FUNCTION_BLOCK basicSensorGenerico (* Logica unica do sensor generico (4-20 mA ou comunicacao) *)
  (* Standard: 61499-2 *)
  (* Version 2.2, 12/11/2026, Hidryco, Hidryco, 2.2: aviso e erro do proprio dispositivo por comunicacao (fldAvisoDisp/fldErroDisp, REQ_FB_DISP): erro diferente de 0 = falha do sensor (cfgTempoFalha); aviso = alarme almAviso; codigos stsCodigoErro/stsCodigoAviso para o diagnostico. 2.1: cfgSkid = sensor sempre habilitado. 2.0: falha do 4-20 mA abaixo de 3800 ou acima de 22000 (eram 3600/21000), confirmada em cfgTempoFalha. 1.9: stsAtivoHH/stsAtivoH (alarme com o tempo do alarme e sem memoria; some quando o valor volta) e stsDisponivel (sensor habilitado, com leitura e sem falha) no CNF. 1.8: limites dos alarmes em unidade de engenharia para o grafico da IHM (stsLimHH..LL; nivel: % x altura maxima / 100). 1.7: stsFalhaSensor (STS_FALHA_SENSOR) so com a falha do sensor (fora da faixa ou falha do instrumento), sem a comunicacao; stsFalhaAtiva e o alarme de falha com qualquer falha. 1.6: IHM: valor, % e bruto no maximo 1 vez por segundo (evento TICK de 1 s); estado, falha e alarmes na hora. 1.5: saida stsFalhaComunicacao (comunicacao do instrumento ou conexao Modbus offline). 1.4: stsFalhaSensor (STS_FALHA_SENSOR na IHM) = falha ativa: sensor em falha agora, sem memoria nem reset; o alarme de falha segue. 1.3: sensor de nivel (cfgNivel) compara os alarmes HH/H/L/LL com a % da altura maxima (setpoints em %); os demais com o valor. 1.2: falha do sinal tambem pelo status da conexao Modbus (fldConexao INT, 1 = online) com cfgUsaConexao, nos dois modos (4-20 mA lido por remota e comunicacao). 1.1: inibicao de L/LL pelo processo e condicao instantanea de cada limite. 1.0: padrao SE.App2CommonProcess - escala, falha NAMUR confirmada por tempo, alarmes HH/H/L/LL com tempo proprio e memoria ate o reset, supressao em falha *)
  PACKAGE Hidryco.HidrycoLib;
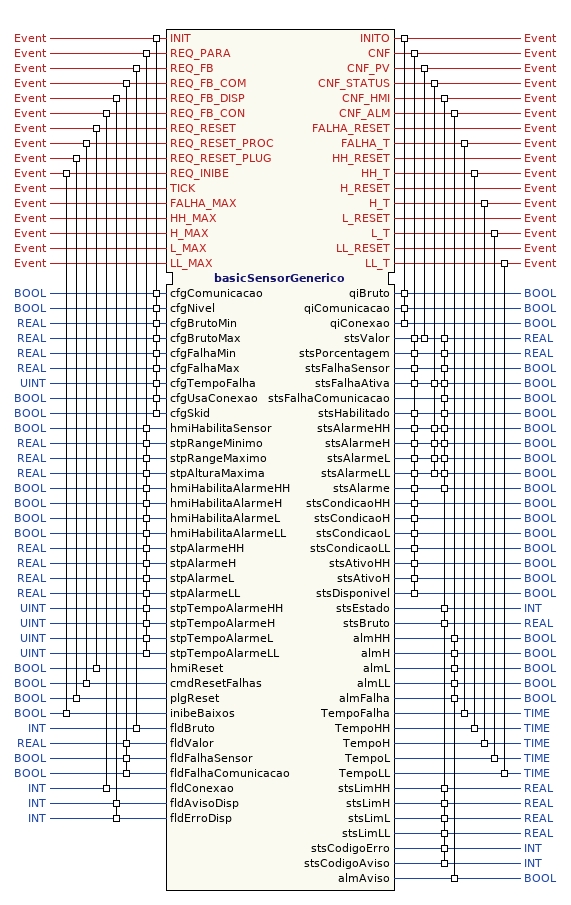
  EVENT_INPUT
    INIT WITH cfgComunicacao, cfgNivel, cfgBrutoMin, cfgBrutoMax, cfgFalhaMin, cfgFalhaMax, cfgTempoFalha, cfgUsaConexao, cfgSkid; (* Inicializacao *)
    REQ_PARA WITH hmiHabilitaSensor, stpRangeMinimo, stpRangeMaximo, stpAlturaMaxima, hmiHabilitaAlarmeHH, hmiHabilitaAlarmeH, hmiHabilitaAlarmeL, hmiHabilitaAlarmeLL, stpAlarmeHH, stpAlarmeH, stpAlarmeL, stpAlarmeLL, stpTempoAlarmeHH, stpTempoAlarmeH, stpTempoAlarmeL, stpTempoAlarmeLL; (* Parametros da IHM (persistentes) *)
    REQ_FB WITH fldBruto; (* Leitura 4-20 mA *)
    REQ_FB_COM WITH fldValor, fldFalhaSensor, fldFalhaComunicacao; (* Leitura por comunicacao *)
    REQ_FB_DISP WITH fldAvisoDisp, fldErroDisp; (* Aviso e erro do proprio dispositivo (comunicacao) *)
    REQ_FB_CON WITH fldConexao; (* Status da conexao Modbus (comunicacao) *)
    REQ_RESET WITH hmiReset; (* Reset pela IHM *)
    REQ_RESET_PROC WITH cmdResetFalhas; (* Reset pelo processo *)
    REQ_RESET_PLUG WITH plgReset; (* Reset pelo plug ISensorStatus *)
    REQ_INIBE WITH inibeBaixos; (* Inibicao dos alarmes L e LL pelo processo *)
    TICK; (* Base de 1 s para atualizar a IHM *)
    FALHA_MAX; (* Fim do tempo de confirmacao da falha (E_DELAY) *)
    HH_MAX; (* Fim do tempo do alarme HH (E_DELAY) *)
    H_MAX; (* Fim do tempo do alarme H (E_DELAY) *)
    L_MAX; (* Fim do tempo do alarme L (E_DELAY) *)
    LL_MAX; (* Fim do tempo do alarme LL (E_DELAY) *)
  END_EVENT
  EVENT_OUTPUT
    INITO WITH qiBruto, qiComunicacao, qiConexao; (* Inicializacao concluida *)
    CNF WITH stsValor, stsPorcentagem, stsFalhaSensor, stsFalhaAtiva, stsHabilitado, stsAlarmeHH, stsAlarmeH, stsAlarmeL, stsAlarmeLL, stsAlarme, stsCondicaoHH, stsCondicaoH, stsCondicaoL, stsCondicaoLL, stsAtivoHH, stsAtivoH, stsDisponivel; (* Status para o processo (na mudanca) *)
    CNF_PV WITH stsValor; (* Valor para o plug (na mudanca) *)
    CNF_STATUS WITH stsAlarmeHH, stsAlarmeH, stsAlarmeL, stsAlarmeLL, stsFalhaAtiva; (* Alarmes para o plug (na mudanca) *)
    CNF_HMI WITH stsValor, stsPorcentagem, stsEstado, stsFalhaSensor, stsFalhaAtiva, stsHabilitado, stsAlarmeHH, stsAlarmeH, stsAlarmeL, stsAlarmeLL, stsAlarme, stsBruto, stsFalhaComunicacao, stsLimHH, stsLimH, stsLimL, stsLimLL, stsCodigoErro, stsCodigoAviso; (* Status para a IHM (na mudanca) *)
    CNF_ALM WITH almHH, almH, almL, almLL, almFalha, almAviso; (* Alarmes para os ALARM_BIT (na mudanca) *)
    FALHA_RESET; (* Cancela o tempo de falha (E_DELAY.STOP) - sai antes do FALHA_T *)
    FALHA_T WITH TempoFalha; (* Inicia o tempo de falha (E_DELAY.START) *)
    HH_RESET; (* Cancela o tempo do alarme HH - sai antes do HH_T *)
    HH_T WITH TempoHH; (* Inicia o tempo do alarme HH *)
    H_RESET; (* Cancela o tempo do alarme H - sai antes do H_T *)
    H_T WITH TempoH; (* Inicia o tempo do alarme H *)
    L_RESET; (* Cancela o tempo do alarme L - sai antes do L_T *)
    L_T WITH TempoL; (* Inicia o tempo do alarme L *)
    LL_RESET; (* Cancela o tempo do alarme LL - sai antes do LL_T *)
    LL_T WITH TempoLL; (* Inicia o tempo do alarme LL *)
  END_EVENT
  VAR_INPUT
    cfgComunicacao : BOOL := FALSE; (* FALSE = entrada 4-20 mA (stsSensorBruto), TRUE = valor por comunicacao (stsEntrada, ja em unidade de engenharia) *)
    cfgNivel : BOOL := FALSE; (* TRUE = sensor de nivel: calcula % sobre a altura maxima *)
    cfgBrutoMin : REAL := 4000.0; (* Valor bruto em 4 mA (TM3: 4000) *)
    cfgBrutoMax : REAL := 20000.0; (* Valor bruto em 20 mA (TM3: 20000) *)
    cfgFalhaMin : REAL := 3800.0; (* Abaixo deste bruto = falha (3,8 mA) *)
    cfgFalhaMax : REAL := 22000.0; (* Acima deste bruto = falha (22,0 mA) *)
    cfgTempoFalha : UINT := 5; (* Tempo para confirmar a falha do sinal (s) *)
    cfgUsaConexao : BOOL := FALSE; (* TRUE = sinal em falha tambem quando o status da conexao Modbus (stsConexao, INT) for diferente de 1 (4-20 mA por remota ou comunicacao) *)
    cfgSkid : BOOL := FALSE; (* TRUE = valor de skid (ja escalado no equipamento): sensor sempre habilitado, sem ajustes na IHM *)
    hmiHabilitaSensor : BOOL; (* IHM: sensor habilitado *)
    stpRangeMinimo : REAL; (* IHM: valor de engenharia em 4 mA *)
    stpRangeMaximo : REAL; (* IHM: valor de engenharia em 20 mA *)
    stpAlturaMaxima : REAL; (* IHM: altura maxima do tanque (nivel) *)
    hmiHabilitaAlarmeHH : BOOL; (* IHM: alarme HH habilitado *)
    hmiHabilitaAlarmeH : BOOL; (* IHM: alarme H habilitado *)
    hmiHabilitaAlarmeL : BOOL; (* IHM: alarme L habilitado *)
    hmiHabilitaAlarmeLL : BOOL; (* IHM: alarme LL habilitado *)
    stpAlarmeHH : REAL; (* IHM: setpoint do alarme HH *)
    stpAlarmeH : REAL; (* IHM: setpoint do alarme H *)
    stpAlarmeL : REAL; (* IHM: setpoint do alarme L *)
    stpAlarmeLL : REAL; (* IHM: setpoint do alarme LL *)
    stpTempoAlarmeHH : UINT; (* IHM: tempo do alarme HH (s) *)
    stpTempoAlarmeH : UINT; (* IHM: tempo do alarme H (s) *)
    stpTempoAlarmeL : UINT; (* IHM: tempo do alarme L (s) *)
    stpTempoAlarmeLL : UINT; (* IHM: tempo do alarme LL (s) *)
    hmiReset : BOOL; (* IHM: reset *)
    cmdResetFalhas : BOOL; (* Processo: reset (com E_RESET_FALHAS) *)
    plgReset : BOOL; (* Plug ISensorStatus: cmdReset *)
    inibeBaixos : BOOL; (* Processo: inibe os alarmes L e LL (ex.: pressao de recalque com as bombas paradas) *)
    fldBruto : INT; (* Campo: valor bruto 4-20 mA *)
    fldValor : REAL; (* Campo (comunicacao): valor em unidade de engenharia *)
    fldFalhaSensor : BOOL; (* Campo (comunicacao): falha do instrumento *)
    fldFalhaComunicacao : BOOL; (* Campo (comunicacao): falha de comunicacao *)
    fldConexao : INT; (* Campo (comunicacao): status da conexao Modbus (connStatusInt: 1 = online, 0 = offline) *)
    fldAvisoDisp : INT; (* Campo (comunicacao): condicao de aviso do proprio dispositivo (0 = nenhum) *)
    fldErroDisp : INT; (* Campo (comunicacao): condicao de erro do proprio dispositivo (0 = nenhum) *)
  END_VAR
  VAR_OUTPUT
    qiBruto : BOOL; (* Assina o symlink 4-20 mA (NOT cfgComunicacao) *)
    qiComunicacao : BOOL; (* Assina os symlinks de comunicacao (cfgComunicacao) *)
    qiConexao : BOOL; (* Assina o symlink do status da conexao (cfgUsaConexao) *)
    stsValor : REAL; (* Valor em unidade de engenharia (0 em falha ou desabilitado) *)
    stsPorcentagem : REAL; (* Nivel em % da altura maxima (so cfgNivel) *)
    stsFalhaSensor : BOOL; (* Falha do sensor (4-20 mA fora da faixa ou falha do instrumento), confirmada e ativa, sem a falha de comunicacao *)
    stsFalhaAtiva : BOOL; (* Qualquer falha confirmada e ativa (sensor ou comunicacao) *)
    stsFalhaComunicacao : BOOL; (* Falha de comunicacao do sensor (falha do instrumento por comunicacao ou conexao Modbus offline) *)
    stsHabilitado : BOOL; (* Sensor habilitado *)
    stsAlarmeHH : BOOL; (* Alarme HH (memorizado ate o reset; suprimido com o sinal em falha) *)
    stsAlarmeH : BOOL; (* Alarme H (memorizado ate o reset; suprimido com o sinal em falha) *)
    stsAlarmeL : BOOL; (* Alarme L (memorizado ate o reset; suprimido com o sinal em falha) *)
    stsAlarmeLL : BOOL; (* Alarme LL (memorizado ate o reset; suprimido com o sinal em falha) *)
    stsAlarme : BOOL; (* Algum alarme ativo *)
    stsCondicaoHH : BOOL; (* Valor alem do setpoint HH agora (sem tempo e sem memoria; so com o alarme habilitado e o sinal bom) *)
    stsCondicaoH : BOOL; (* Valor alem do setpoint H agora (sem tempo e sem memoria; so com o alarme habilitado e o sinal bom) *)
    stsCondicaoL : BOOL; (* Valor alem do setpoint L agora (sem tempo e sem memoria; so com o alarme habilitado e o sinal bom) *)
    stsCondicaoLL : BOOL; (* Valor alem do setpoint LL agora (sem tempo e sem memoria; so com o alarme habilitado e o sinal bom) *)
    stsAtivoHH : BOOL; (* Alarme HH com o tempo do alarme e sem memoria (some quando o valor volta; so com o alarme habilitado e o sinal bom) *)
    stsAtivoH : BOOL; (* Alarme H com o tempo do alarme e sem memoria (some quando o valor volta; so com o alarme habilitado e o sinal bom) *)
    stsDisponivel : BOOL; (* Sensor habilitado, com leitura e sem falha *)
    stsEstado : INT; (* IHM: 0 normal, 1 alerta (H/L), 2 alarme (HH/LL), 3 falha, 4 desabilitado *)
    stsBruto : REAL; (* IHM: valor bruto lido (diagnostico) *)
    almHH : BOOL; (* Entrada do ALARM_BIT HH *)
    almH : BOOL; (* Entrada do ALARM_BIT H *)
    almL : BOOL; (* Entrada do ALARM_BIT L *)
    almLL : BOOL; (* Entrada do ALARM_BIT LL *)
    almFalha : BOOL; (* Entrada do ALARM_BIT de falha do sensor *)
    TempoFalha : TIME; (* E_DELAY da falha *)
    TempoHH : TIME; (* E_DELAY do alarme HH *)
    TempoH : TIME; (* E_DELAY do alarme H *)
    TempoL : TIME; (* E_DELAY do alarme L *)
    TempoLL : TIME; (* E_DELAY do alarme LL *)
    stsLimHH : REAL; (* Limite do alarme HH em unidade de engenharia (para o grafico) *)
    stsLimH : REAL; (* Limite do alarme H em unidade de engenharia (para o grafico) *)
    stsLimL : REAL; (* Limite do alarme L em unidade de engenharia (para o grafico) *)
    stsLimLL : REAL; (* Limite do alarme LL em unidade de engenharia (para o grafico) *)
    stsCodigoErro : INT; (* IHM: codigo de erro do proprio dispositivo (0 = nenhum; diferente de 0 = falha do sensor) *)
    stsCodigoAviso : INT; (* IHM: codigo de aviso do proprio dispositivo (0 = nenhum; so alarme) *)
    almAviso : BOOL; (* Entrada do ALARM_BIT de aviso do proprio dispositivo *)
  END_VAR
  VAR
    initDone : BOOL;
    initPass : BOOL;
    fbRecebido : BOOL; (* Ja houve leitura do campo *)
    bReset : BOOL;
    bRuimAgora : BOOL; (* Sinal fora da faixa / falha agora *)
    bSensorRuim : BOOL; (* Falha do proprio sensor agora (fora da faixa 4-20 mA ou falha do instrumento), sem a comunicacao *)
    bSuprimido : BOOL; (* Alarmes suprimidos *)
    rBruto : REAL;
    rFaixa : REAL;
    rMin : REAL;
    rMax : REAL;
    bTimFalha : BOOL;
    oldTimFalha : BOOL;
    bCondHH : BOOL;
    bMemHH : BOOL;
    bTimHH : BOOL;
    oldTimHH : BOOL;
    bAcimaHH : BOOL;
    bCondH : BOOL;
    bMemH : BOOL;
    bTimH : BOOL;
    oldTimH : BOOL;
    bTempoHH : BOOL; (* Tempo do HH venceu com a condicao presente (sem memoria) *)
    bTempoH : BOOL; (* Tempo do H venceu com a condicao presente (sem memoria) *)
    bAcimaH : BOOL;
    bCondL : BOOL;
    bMemL : BOOL;
    bTimL : BOOL;
    oldTimL : BOOL;
    bAcimaL : BOOL;
    bCondLL : BOOL;
    bMemLL : BOOL;
    bTimLL : BOOL;
    oldTimLL : BOOL;
    bAcimaLL : BOOL;
    oldValor : REAL;
    oldPct : REAL;
    oldBruto : REAL;
    wSts : WORD;
    oldSts : WORD := 16#FFFF;
    wAlm : WORD;
    oldAlm : WORD := 16#FFFF;
    oldCodErro : INT := -1;
    oldCodAviso : INT := -1;
    oldEstado : INT := -1;
    hmiBruto : REAL := -1.0;
    hmiPct : REAL := -1.0;
    hmiValor : REAL := -1.0;
    rCmp : REAL; (* Valor comparado com os alarmes: % (sensor de nivel) ou valor *)
    rEscLim : REAL;
    ostsLimHH : REAL := -1.0;
    ostsLimH : REAL := -1.0;
    ostsLimL : REAL := -1.0;
    ostsLimLL : REAL := -1.0;
  END_VAR
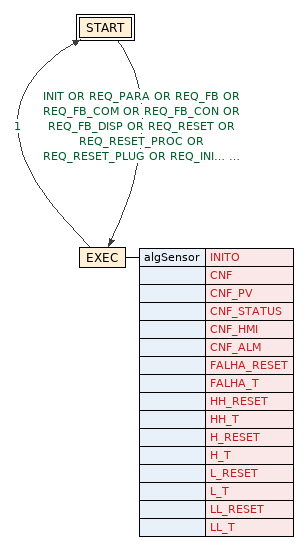
  EC_STATES
    START; (* Estado inicial *)
    EXEC : algSensor -> INITO, -> CNF, -> CNF_PV, -> CNF_STATUS, -> CNF_HMI, -> CNF_ALM, -> FALHA_RESET, -> FALHA_T, -> HH_RESET, -> HH_T, -> H_RESET, -> H_T, -> L_RESET, -> L_T, -> LL_RESET, -> LL_T; (* Executa a logica; o algoritmo decide quais eventos saem *)
  END_STATES
  EC_TRANSITIONS
    START TO EXEC := INIT OR REQ_PARA OR REQ_FB OR REQ_FB_COM OR REQ_FB_CON OR REQ_FB_DISP OR REQ_RESET OR REQ_RESET_PROC OR REQ_RESET_PLUG OR REQ_INIBE OR FALHA_MAX OR HH_MAX OR H_MAX OR L_MAX OR LL_MAX OR TICK;
    EXEC TO START := 1;
  END_TRANSITIONS
  ALGORITHM algSensor IN ST: (* Logica completa do sensor (um unico algoritmo) *)
(* =====================================================================
   basicSensorGenerico v1.1 - logica do CAT Sensor_Generico (HidrycoLib)
   Padrao das bibliotecas Schneider (SE.App2CommonProcess):
   - eventos de saida desligados no inicio e ligados so na mudanca;
   - tempos por E_DELAY externo (X_T / X_RESET / X_MAX), um por alarme;
   - alarmes para o sistema de alarmes do EAE por ALARM_BIT (no CAT).
   Regras (definidas pelo usuario):
   - origem 4-20 mA (escala bruta e limites NAMUR offline) ou comunicacao
     (valor ja em unidade de engenharia);
   - falha do sinal confirmada apos cfgTempoFalha: valor vai a 0 e os
     alarmes ficam suprimidos; a falha vale enquanto o sinal estiver ruim, e o
     sensor volta a funcionar assim que o sinal volta;
   - durante a confirmacao o valor fica congelado (nao vai a 0 por um pico);
   - alarmes HH/H/L/LL sem histerese, cada um com o proprio tempo,
     memorizados ate o reset (IHM, processo ou plug);
   - sensor desabilitado: valor 0, sem falha e sem alarmes.
   v1.3: sensor de nivel (cfgNivel): HH/H/L/LL comparados com a % da altura maxima.
   v1.1: inibeBaixos (processo) inibe L/LL e libera a memoria deles;
         stsCondicaoX = valor alem do setpoint X agora (sem tempo, sem memoria).
   ===================================================================== *)

(* ---- 0. Eventos de saida: so sai o que for ligado abaixo ---- *)
INITO       := FALSE;
CNF         := FALSE;
CNF_PV      := FALSE;
CNF_STATUS  := FALSE;
CNF_HMI     := FALSE;
CNF_ALM     := FALSE;
FALHA_RESET := FALSE;
FALHA_T     := FALSE;
HH_RESET := FALSE; HH_T := FALSE;
H_RESET  := FALSE; H_T  := FALSE;
L_RESET  := FALSE; L_T  := FALSE;
LL_RESET := FALSE; LL_T := FALSE;

IF REQ_FB OR REQ_FB_COM OR REQ_FB_CON THEN
    fbRecebido := TRUE;                    (* campo valido a partir da 1a leitura *)
END_IF;

(* ---- 1. Inicializacao ---- *)
IF INIT THEN
    qiBruto       := NOT cfgComunicacao;   (* so assina o symlink da origem configurada *)
    qiComunicacao := cfgComunicacao;
    qiConexao     := cfgUsaConexao;           (* status da conexao: vale para 4-20 mA lido por remota e para comunicacao *)
    initDone := TRUE;
    initPass := TRUE;
    INITO    := TRUE;
END_IF;
IF NOT initDone THEN
    RETURN;
END_IF;
(* sensor de skid: nao pode ser desabilitado (vale mesmo com FALSE gravado de antes) *)
IF cfgSkid THEN
    hmiHabilitaSensor := TRUE;
END_IF;

(* ---- 2. Sinal ---- *)
IF cfgComunicacao THEN
    rBruto     := fldValor;
    bRuimAgora := fbRecebido AND (fldFalhaSensor OR fldFalhaComunicacao OR (cfgUsaConexao AND fldConexao <> 1));
    bSensorRuim := fbRecebido AND fldFalhaSensor;
ELSE
    rBruto     := INT_TO_REAL(fldBruto);
    bRuimAgora := fbRecebido AND ((rBruto < cfgFalhaMin) OR (rBruto > cfgFalhaMax) OR (cfgUsaConexao AND fldConexao <> 1));
    bSensorRuim := fbRecebido AND ((rBruto < cfgFalhaMin) OR (rBruto > cfgFalhaMax));
END_IF;

(* erro do proprio dispositivo (ex.: SC4500 por Modbus): falha do sensor, confirmada pelo mesmo tempo *)
IF fbRecebido AND (fldErroDisp <> 0) THEN
    bRuimAgora  := TRUE;
    bSensorRuim := TRUE;
END_IF;

(* ---- 3. Falha do sensor: confirmada pelo tempo; vale enquanto o sensor estiver em falha (sem memoria) ---- *)
bReset := (REQ_RESET AND hmiReset) OR (REQ_RESET_PROC AND cmdResetFalhas) OR (REQ_RESET_PLUG AND plgReset);
IF NOT hmiHabilitaSensor THEN
    stsFalhaAtiva := FALSE;
ELSE
    IF FALHA_MAX AND bRuimAgora THEN
        stsFalhaAtiva := TRUE;             (* falha confirmada *)
    END_IF;
    IF NOT bRuimAgora THEN
        stsFalhaAtiva := FALSE;            (* sinal voltou: a falha sai sozinha, sem reset *)
    END_IF;
END_IF;
(* falha de comunicacao (imediata; o tempo de deteccao e o do proprio Modbus) *)
stsFalhaComunicacao := hmiHabilitaSensor AND fbRecebido AND
    ((cfgComunicacao AND fldFalhaComunicacao) OR (cfgUsaConexao AND fldConexao <> 1));
(* STS_FALHA_SENSOR = so a falha do sensor (confirmada pelo tempo); com a comunicacao em falha o valor lido nao vale, entao nao conta *)
stsFalhaSensor := stsFalhaAtiva AND bSensorRuim AND NOT stsFalhaComunicacao;
bTimFalha := hmiHabilitaSensor AND bRuimAgora AND NOT stsFalhaAtiva;
IF bTimFalha <> oldTimFalha THEN
    IF bTimFalha THEN
        TempoFalha := TO_TIME(UINT_TO_DINT(cfgTempoFalha) * 1000);
        FALHA_T := TRUE;
    ELSE
        FALHA_RESET := TRUE;
    END_IF;
    oldTimFalha := bTimFalha;
END_IF;

(* ---- 4. Valor em unidade de engenharia ---- *)
IF NOT hmiHabilitaSensor OR NOT fbRecebido OR stsFalhaAtiva THEN
    stsValor := 0.0;                       (* desabilitado, sem leitura ou falha confirmada *)
ELSIF bRuimAgora THEN
    ;                                      (* confirmando a falha: valor congelado *)
ELSIF cfgComunicacao THEN
    stsValor := fldValor;                  (* ja chega em unidade de engenharia *)
ELSE
    rFaixa := cfgBrutoMax - cfgBrutoMin;
    IF rFaixa <> 0.0 THEN
        stsValor := stpRangeMinimo + (rBruto - cfgBrutoMin) * (stpRangeMaximo - stpRangeMinimo) / rFaixa;
        rMin := MIN(stpRangeMinimo, stpRangeMaximo);
        rMax := MAX(stpRangeMinimo, stpRangeMaximo);
        stsValor := LIMIT(rMin, stsValor, rMax);
    ELSE
        stsValor := 0.0;                   (* escala bruta invalida *)
    END_IF;
END_IF;
IF cfgNivel AND stpAlturaMaxima > 0.0 THEN
    stsPorcentagem := stsValor * 100.0 / stpAlturaMaxima;
ELSE
    stsPorcentagem := 0.0;
END_IF;
stsBruto := rBruto;
(* alarmes do sensor de nivel pela % da altura maxima; os demais pelo valor em unidade de engenharia *)
IF cfgNivel THEN
    rCmp := stsPorcentagem;
ELSE
    rCmp := stsValor;
END_IF;

(* ---- 5. Alarmes (suprimidos com o sensor desabilitado, sem leitura ou em falha) ---- *)
bSuprimido := NOT hmiHabilitaSensor OR NOT fbRecebido OR bRuimAgora OR stsFalhaAtiva;
bAcimaHH := rCmp > stpAlarmeHH;
bCondHH := hmiHabilitaAlarmeHH AND NOT bSuprimido AND bAcimaHH;
stsCondicaoHH := bCondHH;
IF HH_MAX AND bCondHH THEN
    bTempoHH := TRUE;                     (* com tempo, sem memoria *)
    bMemHH := TRUE;                       (* tempo do alarme HH venceu com a condicao presente *)
END_IF;
IF bReset AND NOT bCondHH THEN
    bMemHH := FALSE;                      (* reset so libera se a condicao ja sumiu *)
END_IF;
IF NOT hmiHabilitaAlarmeHH OR NOT hmiHabilitaSensor THEN
    bMemHH := FALSE;                      (* alarme ou sensor desabilitado zera o alarme *)
END_IF;
IF NOT bCondHH THEN
    bTempoHH := FALSE;                    (* condicao sumiu: sai na hora *)
END_IF;
(* o tempo conta a cada vez que a condicao aparece, mesmo com o alarme ainda memorizado (para o stsAtivoHH) *)
bTimHH := bCondHH AND NOT bTempoHH;
IF bTimHH <> oldTimHH THEN
    IF bTimHH THEN
        TempoHH := TO_TIME(UINT_TO_DINT(stpTempoAlarmeHH) * 1000);
        HH_T := TRUE;
    ELSE
        HH_RESET := TRUE;
    END_IF;
    oldTimHH := bTimHH;
END_IF;
stsAlarmeHH := bMemHH AND NOT bSuprimido;
stsAtivoHH := bTempoHH AND bCondHH;

bAcimaH := rCmp > stpAlarmeH;
bCondH := hmiHabilitaAlarmeH AND NOT bSuprimido AND bAcimaH;
stsCondicaoH := bCondH;
IF H_MAX AND bCondH THEN
    bTempoH := TRUE;                     (* com tempo, sem memoria *)
    bMemH := TRUE;                       (* tempo do alarme H venceu com a condicao presente *)
END_IF;
IF bReset AND NOT bCondH THEN
    bMemH := FALSE;                      (* reset so libera se a condicao ja sumiu *)
END_IF;
IF NOT hmiHabilitaAlarmeH OR NOT hmiHabilitaSensor THEN
    bMemH := FALSE;                      (* alarme ou sensor desabilitado zera o alarme *)
END_IF;
IF NOT bCondH THEN
    bTempoH := FALSE;                    (* condicao sumiu: sai na hora *)
END_IF;
(* o tempo conta a cada vez que a condicao aparece, mesmo com o alarme ainda memorizado (para o stsAtivoH) *)
bTimH := bCondH AND NOT bTempoH;
IF bTimH <> oldTimH THEN
    IF bTimH THEN
        TempoH := TO_TIME(UINT_TO_DINT(stpTempoAlarmeH) * 1000);
        H_T := TRUE;
    ELSE
        H_RESET := TRUE;
    END_IF;
    oldTimH := bTimH;
END_IF;
stsAlarmeH := bMemH AND NOT bSuprimido;
stsAtivoH := bTempoH AND bCondH;

bAcimaL := rCmp < stpAlarmeL;
bCondL := hmiHabilitaAlarmeL AND NOT bSuprimido AND bAcimaL AND NOT inibeBaixos;
stsCondicaoL := bCondL;
IF inibeBaixos THEN
    bMemL := FALSE;                      (* inibido pelo processo: libera o que estava memorizado *)
END_IF;
IF L_MAX AND bCondL THEN
    bMemL := TRUE;                       (* tempo do alarme L venceu com a condicao presente *)
END_IF;
IF bReset AND NOT bCondL THEN
    bMemL := FALSE;                      (* reset so libera se a condicao ja sumiu *)
END_IF;
IF NOT hmiHabilitaAlarmeL OR NOT hmiHabilitaSensor THEN
    bMemL := FALSE;                      (* alarme ou sensor desabilitado zera o alarme *)
END_IF;
bTimL := bCondL AND NOT bMemL;
IF bTimL <> oldTimL THEN
    IF bTimL THEN
        TempoL := TO_TIME(UINT_TO_DINT(stpTempoAlarmeL) * 1000);
        L_T := TRUE;
    ELSE
        L_RESET := TRUE;
    END_IF;
    oldTimL := bTimL;
END_IF;
stsAlarmeL := bMemL AND NOT bSuprimido;

bAcimaLL := rCmp < stpAlarmeLL;
bCondLL := hmiHabilitaAlarmeLL AND NOT bSuprimido AND bAcimaLL AND NOT inibeBaixos;
stsCondicaoLL := bCondLL;
IF inibeBaixos THEN
    bMemLL := FALSE;                      (* inibido pelo processo: libera o que estava memorizado *)
END_IF;
IF LL_MAX AND bCondLL THEN
    bMemLL := TRUE;                       (* tempo do alarme LL venceu com a condicao presente *)
END_IF;
IF bReset AND NOT bCondLL THEN
    bMemLL := FALSE;                      (* reset so libera se a condicao ja sumiu *)
END_IF;
IF NOT hmiHabilitaAlarmeLL OR NOT hmiHabilitaSensor THEN
    bMemLL := FALSE;                      (* alarme ou sensor desabilitado zera o alarme *)
END_IF;
bTimLL := bCondLL AND NOT bMemLL;
IF bTimLL <> oldTimLL THEN
    IF bTimLL THEN
        TempoLL := TO_TIME(UINT_TO_DINT(stpTempoAlarmeLL) * 1000);
        LL_T := TRUE;
    ELSE
        LL_RESET := TRUE;
    END_IF;
    oldTimLL := bTimLL;
END_IF;
stsAlarmeLL := bMemLL AND NOT bSuprimido;

stsAlarme := stsAlarmeHH OR stsAlarmeH OR stsAlarmeL OR stsAlarmeLL;
stsHabilitado := hmiHabilitaSensor;
stsDisponivel := hmiHabilitaSensor AND fbRecebido AND NOT bRuimAgora AND NOT stsFalhaAtiva;

(* ---- 6. Entradas dos ALARM_BIT (lista de alarmes do EAE) ---- *)
almHH := stsAlarmeHH;
almH  := stsAlarmeH;
almL  := stsAlarmeL;
almLL := stsAlarmeLL;
almFalha := stsFalhaAtiva;                (* alarme de falha: sensor ou comunicacao *)

(* ---- 7. Estado para o simbolo ---- *)
IF NOT hmiHabilitaSensor THEN
    stsEstado := 4;
ELSIF stsFalhaSensor OR stsFalhaAtiva THEN
    stsEstado := 3;
ELSIF stsAlarmeHH OR stsAlarmeLL THEN
    stsEstado := 2;
ELSIF stsAlarmeH OR stsAlarmeL THEN
    stsEstado := 1;
ELSE
    stsEstado := 0;
END_IF;

(* ---- 8. Eventos so na mudanca ---- *)
wSts := 0;
IF stsFalhaSensor THEN wSts := wSts OR 16#0001; END_IF;
IF stsFalhaAtiva  THEN wSts := wSts OR 16#0002; END_IF;
IF stsHabilitado  THEN wSts := wSts OR 16#0004; END_IF;
IF stsAlarmeHH    THEN wSts := wSts OR 16#0010; END_IF;
IF stsAlarmeH     THEN wSts := wSts OR 16#0020; END_IF;
IF stsAlarmeL     THEN wSts := wSts OR 16#0040; END_IF;
IF stsAlarmeLL    THEN wSts := wSts OR 16#0080; END_IF;
IF stsCondicaoHH  THEN wSts := wSts OR 16#0100; END_IF;
IF stsCondicaoH   THEN wSts := wSts OR 16#0200; END_IF;
IF stsCondicaoL   THEN wSts := wSts OR 16#0400; END_IF;
IF stsCondicaoLL  THEN wSts := wSts OR 16#0800; END_IF;
IF stsFalhaComunicacao THEN wSts := wSts OR 16#1000; END_IF;
IF stsAtivoHH    THEN wSts := wSts OR 16#2000; END_IF;
IF stsAtivoH     THEN wSts := wSts OR 16#4000; END_IF;
IF stsDisponivel THEN wSts := wSts OR 16#8000; END_IF;
(* codigos do proprio dispositivo para o diagnostico; aviso = so alarme *)
IF hmiHabilitaSensor THEN
    stsCodigoErro  := fldErroDisp;
    stsCodigoAviso := fldAvisoDisp;
ELSE
    stsCodigoErro  := 0;
    stsCodigoAviso := 0;
END_IF;
almAviso := hmiHabilitaSensor AND fbRecebido AND (fldAvisoDisp <> 0) AND NOT stsFalhaComunicacao;
wAlm := 0;
IF almHH    THEN wAlm := wAlm OR 16#0001; END_IF;
IF almH     THEN wAlm := wAlm OR 16#0002; END_IF;
IF almL     THEN wAlm := wAlm OR 16#0004; END_IF;
IF almLL    THEN wAlm := wAlm OR 16#0008; END_IF;
IF almFalha THEN wAlm := wAlm OR 16#0010; END_IF;
IF almAviso THEN wAlm := wAlm OR 16#0020; END_IF;

(* limites dos alarmes em unidade de engenharia (grafico da IHM); nivel: setpoints em % da altura maxima *)
IF cfgNivel THEN
    rEscLim := stpAlturaMaxima / 100.0;
ELSE
    rEscLim := 1.0;
END_IF;
stsLimHH := stpAlarmeHH * rEscLim;
stsLimH  := stpAlarmeH * rEscLim;
stsLimL  := stpAlarmeL * rEscLim;
stsLimLL := stpAlarmeLL * rEscLim;

CNF_PV     := initPass OR (stsValor <> oldValor);
CNF_STATUS := initPass OR ((wSts AND 16#00F2) <> (oldSts AND 16#00F2));
CNF        := initPass OR (stsValor <> oldValor) OR (stsPorcentagem <> oldPct) OR (wSts <> oldSts);
(* IHM: estado/falha/alarme na hora; valor, % e bruto no maximo 1 vez por segundo (TICK) *)
CNF_HMI    := initPass OR (wSts <> oldSts) OR (stsEstado <> oldEstado) OR (stsCodigoErro <> oldCodErro) OR (stsCodigoAviso <> oldCodAviso)
              OR (TICK AND ((stsValor <> hmiValor) OR (stsPorcentagem <> hmiPct) OR (rBruto <> hmiBruto)))
              OR (stsLimHH <> ostsLimHH) OR (stsLimH <> ostsLimH) OR (stsLimL <> ostsLimL) OR (stsLimLL <> ostsLimLL);
IF CNF_HMI THEN
    hmiValor := stsValor; hmiPct := stsPorcentagem; hmiBruto := rBruto;
    ostsLimHH := stsLimHH; ostsLimH := stsLimH; ostsLimL := stsLimL; ostsLimLL := stsLimLL;
END_IF;
CNF_ALM    := initPass OR (wAlm <> oldAlm);
oldValor  := stsValor;
oldPct    := stsPorcentagem;
oldBruto  := rBruto;
oldSts    := wSts;
oldAlm    := wAlm;
oldEstado := stsEstado;
oldCodErro  := stsCodigoErro;
oldCodAviso := stsCodigoAviso;

initPass := FALSE;
  END_ALGORITHM
END_FUNCTION_BLOCK
